(* IEC 61131-3 sources: station-control-three-platforms/codesys/src (part 2) *)

(* ---- GVL_TestResult.st ---- *)
// Result of the test bench (FB_TestBench). Port of DB_TestResult; read by codesys/scripts/build_and_run.py.
{attribute 'qualified_only'}
VAR_GLOBAL
    Done : BOOL;   // the bench has finished; the values below no longer change
    AllPassed : BOOL;   // Done and every case passed
    CasesTotal : INT;
    CasesRun : INT;
    CasesPassed : INT;
    CasesFailed : INT;
    FirstFailedCase : INT;   // 0 = none
    FirstFailedCheck : INT;   // 0 = none; codes in the header of FB_TestBench
    MaxFeatError : REAL;   // N or mm, largest difference of an element from its expected value
    BenchCalls : DINT;   // task cycles the bench needed
    CasePass : ARRAY[1..32] OF BOOL;
    CaseCheck : ARRAY[1..32] OF INT;   // failed check of each case, 0 = passed
    CaseNok : ARRAY[1..32] OF INT;   // NOK code the block gave in each case
END_VAR

(* ---- FB_CurveEval.st ---- *)
FUNCTION_BLOCK FB_CurveEval
//  CODESYS V3.5 port of the Siemens SCL block. Only the syntax changed: no # before local names,
//  REGION as {region} pragma, global data as qualified GVL names, LIMIT with positional arguments.
//  Called in the cyclic interrupt that samples the load cell and the axis position.
//  Nothing is stored as a curve: every evaluation element is updated with the new sample.
//  The block works on static variables and writes its outputs once, at the end of every call.
//  Elements (DOSSIER section 6.3):
//    gate 1 (GateX)    pull force FpG1 and return force FrG1 at the same travel;
//                      FMean = (FpG1 + FrG1) / 2 is the spring, FHyst = FpG1 - FrG1 is twice the friction
//    gate 2 (Gate2X)   pull force after the cable is taut
//    peak window       highest pull force between PeakXLo and PeakXHi and its travel (latch release)
//    step              force drop within StepSpan after the peak
//    stop              travel at which the pull force crosses StopF (end stop)
//    envelope          pull force at fixed travel nodes against EnvLo / EnvHi
//  Mode: 1 peak force only, 2 pull-stroke windows, 3 windows with return stroke, 4 envelope.
//  NokCode: 0 OK, 1 element not measured, 2 gate-1 force (spring), 3 hysteresis (friction),
//           4 no return force, 5 gate-2 force, 6 peak force, 7 peak travel, 8 release step,
//           9 stop travel, 10 envelope.
   VAR_INPUT
      Reset : Bool;   // clear all results, before a new pull
      Sample : Bool;   // X and F are a new sample
      Stroke : Int;   // 1 pull, 2 return
      X : Real;   // mm, travel from touch
      F : Real;   // N
      Finish : Bool;   // return stroke finished: judge
      Mode : Int := 3;
      GateX : Real := 3.0;   // mm
      Gate2X : Real := 10.0;   // mm
      PeakXLo : Real := 13.0;   // mm
      PeakXHi : Real := 26.0;   // mm
      StepSpan : Real := 2.0;   // mm
      StopF : Real := 30.0;   // N
      G1Lo : Real;   // N, limits of FpG1 (mode 2)
      G1Hi : Real;
      MeanLo : Real;   // N, limits of FMean (mode 3)
      MeanHi : Real;
      HystLo : Real;   // N, limits of FHyst (mode 3)
      HystHi : Real;
      RetFMin : Real;   // N, FrG1 must be above (mode 3)
      G2Lo : Real;   // N, limits of FpG2
      G2Hi : Real;
      PeakFLo : Real;   // N
      PeakFHi : Real;
      PeakXMin : Real;   // mm, limits of XPeak
      PeakXMax : Real;
      StepLo : Real;   // N
      StopXLo : Real;   // mm
      StopXHi : Real;
      EnvX0 : Real := 1.0;   // mm, first envelope node
      EnvDx : Real := 0.5;   // mm, node spacing
      EnvN : Int := 55;   // number of nodes, at most 64
      EnvLo : Array[0..63] of Real;   // N
      EnvHi : Array[0..63] of Real;   // N
   END_VAR

   VAR_OUTPUT
      FpG1 : Real;
      FrG1 : Real;
      FMean : Real;
      FHyst : Real;
      FpG2 : Real;
      FPeak : Real;
      XPeak : Real;
      FStep : Real;
      XStop : Real;
      EnvViol : Int;   // envelope nodes outside the band
      EnvNodes : Int;   // envelope nodes evaluated
      NSamples : Int;
      Done : Bool;
      Ok : Bool;
      NokCode : Int;
   END_VAR

   VAR
      sHavePrev : Bool;
      sPrevX : Real;
      sPrevF : Real;
      sPrevStroke : Int;
      sGotG1 : Bool;
      sGotG2 : Bool;
      sGotR1 : Bool;
      sGotPeak : Bool;
      sGotStop : Bool;
      sFMin : Real;
      sFpG1 : Real;
      sFrG1 : Real;
      sFMean : Real;
      sFHyst : Real;
      sFpG2 : Real;
      sFPeak : Real;
      sXPeak : Real;
      sFStep : Real;
      sXStop : Real;
      sEnvViol : Int;
      sEnvNodes : Int;
      sNSamples : Int;
      sDone : Bool;
      sOk : Bool;
      sNokCode : Int;
   END_VAR

   VAR_TEMP
      tI : Int;
      tNodeX : Real;
      tFn : Real;
      tCode : Int;
   END_VAR

(* @IMPLEMENTATION *)
    {region "Reset"}
        IF Reset THEN
            sFpG1 := 0.0;
            sFrG1 := 0.0;
            sFMean := 0.0;
            sFHyst := 0.0;
            sFpG2 := 0.0;
            sFPeak := 0.0;
            sXPeak := 0.0;
            sFStep := 0.0;
            sXStop := 0.0;
            sEnvViol := 0;
            sEnvNodes := 0;
            sNSamples := 0;
            sDone := FALSE;
            sOk := FALSE;
            sNokCode := 0;
            sHavePrev := FALSE;
            sGotG1 := FALSE;
            sGotG2 := FALSE;
            sGotR1 := FALSE;
            sGotPeak := FALSE;
            sGotStop := FALSE;
            sFMin := 0.0;
        END_IF;
    {endregion}

    {region "PullStroke"}
        IF NOT Reset AND Sample AND NOT sDone AND Stroke = 1 THEN
            IF sHavePrev AND sPrevStroke = 1 THEN
                // gates: force at a set travel, linear between the two samples around it
                IF NOT sGotG1 AND sPrevX < GateX AND X >= GateX THEN
                    sFpG1 := sPrevF + (F - sPrevF) * (GateX - sPrevX) / (X - sPrevX);
                    sGotG1 := TRUE;
                END_IF;
                IF NOT sGotG2 AND sPrevX < Gate2X AND X >= Gate2X THEN
                    sFpG2 := sPrevF + (F - sPrevF) * (Gate2X - sPrevX) / (X - sPrevX);
                    sGotG2 := TRUE;
                END_IF;
                // end stop: travel at a set force
                IF NOT sGotStop AND sPrevX > Gate2X AND sPrevF < StopF AND F >= StopF THEN
                    sXStop := sPrevX + (X - sPrevX) * (StopF - sPrevF) / (F - sPrevF);
                    sGotStop := TRUE;
                END_IF;
                // envelope: at most four nodes can lie between two samples
                FOR tI := 1 TO 4 DO
                    tNodeX := EnvX0 + EnvDx * INT_TO_REAL(sEnvNodes);
                    IF sEnvNodes < EnvN AND sPrevX < tNodeX AND X >= tNodeX THEN
                        tFn := sPrevF + (F - sPrevF) * (tNodeX - sPrevX) / (X - sPrevX);
                        IF tFn < EnvLo[sEnvNodes] OR tFn > EnvHi[sEnvNodes] THEN
                            sEnvViol := sEnvViol + 1;
                        END_IF;
                        sEnvNodes := sEnvNodes + 1;
                    END_IF;
                END_FOR;
            END_IF;
            // latch release: peak inside the window, then the drop after it
            IF X >= PeakXLo AND X <= PeakXHi AND (NOT sGotPeak OR F > sFPeak) THEN
                sFPeak := F;
                sXPeak := X;
                sFMin := F;
                sGotPeak := TRUE;
            ELSIF sGotPeak AND X <= sXPeak + StepSpan AND F < sFMin THEN
                sFMin := F;
            END_IF;
            IF sGotPeak THEN
                sFStep := sFPeak - sFMin;
            END_IF;
        END_IF;
    {endregion}

    {region "ReturnStroke"}
        IF NOT Reset AND Sample AND NOT sDone AND Stroke = 2 AND sHavePrev THEN
            IF NOT sGotR1 AND sPrevX > GateX AND X <= GateX THEN
                sFrG1 := sPrevF + (F - sPrevF) * (GateX - sPrevX) / (X - sPrevX);
                sGotR1 := TRUE;
            END_IF;
        END_IF;
    {endregion}

    {region "Bookkeeping"}
        IF NOT Reset AND Sample AND NOT sDone THEN
            sPrevX := X;
            sPrevF := F;
            sPrevStroke := Stroke;
            sHavePrev := TRUE;
            IF sNSamples < 32000 THEN
                sNSamples := sNSamples + 1;
            END_IF;
        END_IF;
    {endregion}

    {region "Verdict"}
        IF NOT Reset AND Finish AND NOT sDone THEN
            sFMean := (sFpG1 + sFrG1) * 0.5;
            sFHyst := sFpG1 - sFrG1;
            tCode := 0;
            CASE Mode OF
                1:  // peak force only
                    IF NOT sGotPeak THEN
                        tCode := 1;
                    ELSIF sFPeak < PeakFLo OR sFPeak > PeakFHi THEN
                        tCode := 6;
                    END_IF;
                2, 3:  // windows; mode 3 judges gate 1 with the return stroke
                    IF NOT (sGotG1 AND sGotG2 AND sGotPeak AND sGotStop) THEN
                        tCode := 1;
                    ELSIF Mode = 3 AND NOT sGotR1 THEN
                        tCode := 1;
                    ELSIF Mode = 2 AND (sFpG1 < G1Lo OR sFpG1 > G1Hi) THEN
                        tCode := 2;
                    ELSIF Mode = 3 AND (sFMean < MeanLo OR sFMean > MeanHi) THEN
                        tCode := 2;
                    ELSIF Mode = 3 AND (sFHyst < HystLo OR sFHyst > HystHi) THEN
                        tCode := 3;
                    ELSIF Mode = 3 AND sFrG1 < RetFMin THEN
                        tCode := 4;
                    ELSIF sFpG2 < G2Lo OR sFpG2 > G2Hi THEN
                        tCode := 5;
                    ELSIF sFPeak < PeakFLo OR sFPeak > PeakFHi THEN
                        tCode := 6;
                    ELSIF sXPeak < PeakXMin OR sXPeak > PeakXMax THEN
                        tCode := 7;
                    ELSIF sFStep < StepLo THEN
                        tCode := 8;
                    ELSIF sXStop < StopXLo OR sXStop > StopXHi THEN
                        tCode := 9;
                    END_IF;
                4:  // envelope: every node reached and inside
                    IF sEnvNodes < EnvN THEN
                        tCode := 1;
                    ELSIF sEnvViol > 0 THEN
                        tCode := 10;
                    END_IF;
                ELSE
                    tCode := 1;
            END_CASE;
            sNokCode := tCode;
            sOk := tCode = 0;
            sDone := TRUE;
        END_IF;
    {endregion}

    {region "Outputs"}
        // the working values live in static variables; the outputs are written here and nowhere else
        FpG1 := sFpG1;
        FrG1 := sFrG1;
        FMean := sFMean;
        FHyst := sFHyst;
        FpG2 := sFpG2;
        FPeak := sFPeak;
        XPeak := sXPeak;
        FStep := sFStep;
        XStop := sXStop;
        EnvViol := sEnvViol;
        EnvNodes := sEnvNodes;
        NSamples := sNSamples;
        Done := sDone;
        Ok := sOk;
        NokCode := sNokCode;
    {endregion}
END_FUNCTION_BLOCK

(* ---- FB_HandleStation.st ---- *)
FUNCTION_BLOCK FB_HandleStation
//  CODESYS V3.5 port of the Siemens SCL block (siemens/scl/FB_HandleStation.scl). Changes, all forced
//  by the compiler: the timer variable sT is sTim (ST is a keyword, identifiers are not case-sensitive);
//  the evaluation recipe comes in by reference (Rcp) and is copied into Eval at the tare, because the
//  caller may not write into Eval from outside (C0037).
//  Called in the same cyclic interrupt as the sampling (CycleTime).
//  States (DOSSIER section 3):
//    0 Idle         wait for a part; check presence time and the LH/RH sensor pattern
//    1 Clamp        close the clamp
//    2 Tare         zero the load cell with the hook free
//    3 Approach     drive towards the grip until the force passes FTouch; the touch position
//                   must lie in its window
//    4 Pull         sample every cycle into the curve evaluation; reverse at FRev
//    5 Return       sample the return stroke down to travel 0, then go home fast
//    6 Evaluate     judge
//    7 UnloadOk     open the clamp; wait until the part has left
//    8 RejectLock   open the clamp; the station stays locked until the part has left AND the
//                   reject-chute sensor has seen a part pass
//    9 Fault        drive stopped; after the acknowledge the axis goes home and the part that was
//                   in test is treated as rejected (an interrupted test is not a passed test)
//   10 Home         go home after a fault
//  NokCode: 1 to 10 from FB_CurveEval; 20 wrong hand or sensor pattern not plausible;
//           21 no touch or touch outside its window; 22 force above FAbsMax; 23 no end stop;
//           24 test interrupted by a fault.
//  FaultCode: 1 safety circuit open, 2 drive not ready, 3 clamp time-out, 4 load cell does not tare.
   VAR_INPUT
      CycleTime : Real := 0.002;   // s
      SafetyOk : Bool;
      DriveOk : Bool;
      AckFault : Bool;
      StartEnable : Bool;   // release from the line
      PartPresent : Bool;
      SensLH : Bool;   // variant sensor that only an LH unit covers
      SensRH : Bool;   // variant sensor that only an RH unit covers
      VariantLH : Bool;   // recipe: TRUE = LH units are being built
      ClampClosed : Bool;
      ClampOpen : Bool;
      RejectChute : Bool;   // light barrier in the reject chute
      Pos : Real;   // mm, axis position, 0 = home
      Force : Real;   // N, load cell
      VPull : Real := 50.0;   // mm/s
      VHome : Real := 150.0;   // mm/s
      FTouch : Real := 1.5;   // N
      FRev : Real := 40.0;   // N
      FAbsMax : Real := 60.0;   // N, protects the painted part
      XMax : Real := 38.0;   // mm
      TouchLo : Real := 3.0;   // mm, window of the touch position
      TouchHi : Real := 7.0;
      Compliance : Real := 0.025;   // mm/N, rig deflection taken out of the travel
      TareTol : Real := 0.5;   // N
      TPresent : Real := 0.1;   // s
      TClampMax : Real := 1.0;   // s
      TRejectWarn : Real := 30.0;   // s
      MaxConsecNok : Int := 3;
   END_VAR

   VAR_IN_OUT
      Rcp : ST_EvalRecipe;   // evaluation recipe, copied into Eval at every tare
   END_VAR

   VAR_OUTPUT
      QClamp : Bool;
      QDriveEnable : Bool;
      QVel : Real;   // mm/s, positive = pull
      QLampOk : Bool;
      QLampNok : Bool;
      QCallOperator : Bool;
      State : Int;
      Verdict : Int;   // 0 none, 1 OK, 2 NOK
      NokCode : Int;
      FaultCode : Int;
      Locked : Bool;
      RigCheckRequired : Bool;   // too many rejects in a row: run the master part
      XTravel : Real;   // mm
      FNet : Real;   // N
      TCycle : Real;   // s, clamp to verdict of the last part
      CntTotal : DInt;
      CntOk : DInt;
      CntNok : DInt;
      CntRejectConfirmed : DInt;
      CntConsecNok : Int;
      CntByCode : Array[0..31] of DInt;
   END_VAR

   VAR
      Eval : FB_CurveEval;
      sTim : Real;
      sTCycle : Real;
      sTare : Real;
      sTouchPos : Real;
      sFTouch : Real;
      sPreNok : Int;
      sPartGone : Bool;
      sChutePrev : Bool;
      sInTest : Bool;
      sWasLocked : Bool;
      sState : Int;
      sRigCheckRequired : Bool;
      sCntTotal : DInt;
      sCntOk : DInt;
      sCntNok : DInt;
      sCntRejectConfirmed : DInt;
      sCntConsecNok : Int;
      sCntByCode : Array[0..31] of DInt;
   END_VAR

   VAR_TEMP
      tVariantOk : Bool;
      tChuteEdge : Bool;
      tCode : Int;
   END_VAR

(* @IMPLEMENTATION *)
    {region "Inputs"}
        FNet := Force - sTare;
        tChuteEdge := RejectChute AND NOT sChutePrev;
        sChutePrev := RejectChute;
        sTim := sTim + CycleTime;
        sTCycle := sTCycle + CycleTime;
        QVel := 0.0;
        // exactly the sensor of the expected hand, and not the other one
        tVariantOk := (VariantLH AND SensLH AND NOT SensRH) OR (NOT VariantLH AND SensRH AND NOT SensLH);
    {endregion}

    {region "Faults"}
        IF sState <> 9 AND (NOT SafetyOk OR NOT DriveOk) THEN
            IF NOT SafetyOk THEN
                FaultCode := 1;
            ELSE
                FaultCode := 2;
            END_IF;
            IF sState <> 10 THEN
                sInTest := sState >= 1 AND sState <= 6;
                sWasLocked := sState = 8;
            END_IF;
            sState := 9;
        END_IF;
    {endregion}

    {region "Sequence"}
        CASE sState OF
            0:  // Idle
                Locked := FALSE;
                IF NOT PartPresent THEN
                    sTim := 0.0;
                    QLampOk := FALSE;
                    QLampNok := FALSE;
                ELSIF sTim >= TPresent AND StartEnable AND ClampOpen AND NOT sRigCheckRequired THEN
                    Verdict := 0;
                    NokCode := 0;
                    sPreNok := 0;
                    sTCycle := 0.0;
                    sTim := 0.0;
                    IF tVariantOk THEN
                        sState := 1;
                    ELSE
                        sPreNok := 20;   // never pull a part of the wrong hand
                        sState := 6;
                    END_IF;
                END_IF;
            1:  // Clamp
                QClamp := TRUE;
                IF ClampClosed THEN
                    sTim := 0.0;
                    sState := 2;
                ELSIF sTim > TClampMax THEN
                    FaultCode := 3;
                    sInTest := TRUE;
                    sState := 9;
                END_IF;
            2:  // Tare
                IF sTim >= 0.05 THEN
                    IF ABS(Force) > TareTol THEN
                        FaultCode := 4;
                        sInTest := TRUE;
                        sState := 9;
                    ELSE
                        sTare := Force;
                        // the recipe of this part (Siemens: written into Eval by the caller)
                        Eval.Mode := Rcp.Mode;
                        Eval.GateX := Rcp.GateX;
                        Eval.Gate2X := Rcp.Gate2X;
                        Eval.PeakXLo := Rcp.PeakXLo;
                        Eval.PeakXHi := Rcp.PeakXHi;
                        Eval.StepSpan := Rcp.StepSpan;
                        Eval.StopF := Rcp.StopF;
                        Eval.G1Lo := Rcp.G1Lo;
                        Eval.G1Hi := Rcp.G1Hi;
                        Eval.MeanLo := Rcp.MeanLo;
                        Eval.MeanHi := Rcp.MeanHi;
                        Eval.HystLo := Rcp.HystLo;
                        Eval.HystHi := Rcp.HystHi;
                        Eval.RetFMin := Rcp.RetFMin;
                        Eval.G2Lo := Rcp.G2Lo;
                        Eval.G2Hi := Rcp.G2Hi;
                        Eval.PeakFLo := Rcp.PeakFLo;
                        Eval.PeakFHi := Rcp.PeakFHi;
                        Eval.PeakXMin := Rcp.PeakXMin;
                        Eval.PeakXMax := Rcp.PeakXMax;
                        Eval.StepLo := Rcp.StepLo;
                        Eval.StopXLo := Rcp.StopXLo;
                        Eval.StopXHi := Rcp.StopXHi;
                        Eval.EnvX0 := Rcp.EnvX0;
                        Eval.EnvDx := Rcp.EnvDx;
                        Eval.EnvN := Rcp.EnvN;
                        Eval.EnvLo := Rcp.EnvLo;
                        Eval.EnvHi := Rcp.EnvHi;
                        Eval(Reset := TRUE, Sample := FALSE, Stroke := 0, X := 0.0, F := 0.0, Finish := FALSE);
                        sState := 3;
                    END_IF;
                END_IF;
            3:  // Approach
                QVel := VPull;
                IF FNet > FTouch THEN
                    sTouchPos := Pos;
                    sFTouch := FNet;
                    IF Pos < TouchLo OR Pos > TouchHi THEN
                        sPreNok := 21;
                        sState := 5;
                    ELSE
                        XTravel := 0.0;
                        Eval(Reset := FALSE, Sample := TRUE, Stroke := 1, X := 0.0, F := FNet, Finish := FALSE);
                        sState := 4;
                    END_IF;
                ELSIF Pos > TouchHi THEN
                    sPreNok := 21;
                    sTouchPos := Pos;
                    sFTouch := 0.0;
                    sState := 5;
                END_IF;
            4:  // Pull
                QVel := VPull;
                XTravel := Pos - sTouchPos - (FNet - sFTouch) * Compliance;
                Eval(Reset := FALSE, Sample := TRUE, Stroke := 1, X := XTravel, F := FNet, Finish := FALSE);
                IF FNet >= FAbsMax THEN
                    sPreNok := 22;
                    sState := 5;
                ELSIF FNet >= FRev THEN
                    sState := 5;
                ELSIF XTravel >= XMax THEN
                    sPreNok := 23;
                    sState := 5;
                END_IF;
            5:  // Return
                XTravel := Pos - sTouchPos - (FNet - sFTouch) * Compliance;
                IF Pos > sTouchPos - 0.5 THEN
                    QVel := -VPull;
                    IF sPreNok = 0 THEN
                        Eval(Reset := FALSE, Sample := TRUE, Stroke := 2, X := XTravel, F := FNet, Finish := FALSE);
                    END_IF;
                ELSIF Pos > 0.05 THEN
                    QVel := -VHome;
                ELSE
                    sState := 6;
                END_IF;
            6:  // Evaluate
                IF sPreNok <> 0 THEN
                    tCode := sPreNok;
                ELSE
                    Eval(Reset := FALSE, Sample := FALSE, Stroke := 0, X := 0.0, F := 0.0, Finish := TRUE);
                    tCode := Eval.NokCode;
                END_IF;
                NokCode := tCode;
                TCycle := sTCycle;
                sCntTotal := sCntTotal + 1;
                sCntByCode[tCode] := sCntByCode[tCode] + 1;
                QClamp := FALSE;
                sTim := 0.0;
                IF tCode = 0 THEN
                    Verdict := 1;
                    sCntOk := sCntOk + 1;
                    sCntConsecNok := 0;
                    QLampOk := TRUE;
                    sState := 7;
                ELSE
                    Verdict := 2;
                    sCntNok := sCntNok + 1;
                    sCntConsecNok := sCntConsecNok + 1;
                    QLampNok := TRUE;
                    sPartGone := FALSE;
                    sState := 8;
                END_IF;
            7:  // UnloadOk
                QClamp := FALSE;
                IF NOT PartPresent AND ClampOpen THEN
                    sTim := 0.0;
                    sState := 0;
                END_IF;
            8:  // RejectLock
                QClamp := FALSE;
                Locked := TRUE;
                IF NOT PartPresent THEN
                    sPartGone := TRUE;
                END_IF;
                QCallOperator := sTim > TRejectWarn OR sRigCheckRequired;
                IF sPartGone AND tChuteEdge THEN
                    sCntRejectConfirmed := sCntRejectConfirmed + 1;
                    sRigCheckRequired := sCntConsecNok >= MaxConsecNok;
                    QCallOperator := sRigCheckRequired;
                    Locked := FALSE;
                    sTim := 0.0;
                    sState := 0;
                END_IF;
            9:  // Fault
                QClamp := sInTest;
                QCallOperator := TRUE;
                IF AckFault AND SafetyOk AND DriveOk THEN
                    FaultCode := 0;
                    QCallOperator := FALSE;
                    sState := 10;
                END_IF;
            10:  // Home
                IF Pos > 0.05 THEN
                    QVel := -VPull;
                ELSIF sInTest THEN
                    sInTest := FALSE;
                    sPreNok := 24;
                    sState := 6;
                ELSIF sWasLocked THEN
                    sWasLocked := FALSE;   // a fault does not release the reject lock
                    sState := 8;
                ELSE
                    sState := 0;
                END_IF;
            ELSE
                sState := 9;
        END_CASE;
    {endregion}

    {region "RigCheck"}
        // the lock after too many rejects in a row is released by the acknowledge key
        IF sRigCheckRequired AND AckFault AND sState = 0 THEN
            sRigCheckRequired := FALSE;
            sCntConsecNok := 0;
            QCallOperator := FALSE;
        END_IF;
        QDriveEnable := SafetyOk AND DriveOk AND sState <> 9;
    {endregion}

    {region "Outputs"}
        // state and counters live in static variables; these outputs are written here and nowhere else
        State := sState;
        RigCheckRequired := sRigCheckRequired;
        CntTotal := sCntTotal;
        CntOk := sCntOk;
        CntNok := sCntNok;
        CntRejectConfirmed := sCntRejectConfirmed;
        CntConsecNok := sCntConsecNok;
        CntByCode := sCntByCode;
    {endregion}
END_FUNCTION_BLOCK

(* ---- FB_TestBench.st ---- *)
FUNCTION_BLOCK FB_TestBench
//  CODESYS V3.5 port of siemens/scl/test/FB_TestBench.scl. Changes: sT is sTim; the station recipe is
//  the local structure StationRcp, passed to the station as Rcp (Siemens: Station.Eval.* written directly).
//  Called from OB1 every cycle. Needs no input from outside. Finishes on its own, then holds its
//  result in DB_TestResult.
//  Part 1, replay cases 1..NCases (DB_TestData): a recorded curve goes sample by sample into
//    FB_CurveEval. Verdict, NOK code, the nine elements and the envelope counts must equal the
//    values the NumPy evaluation gave for the same samples (elements within DB_TestData.Tol).
//  Part 2, six station cases: FB_HandleStation runs against FB_TestPlant.
//    NCases+1  good LH unit is clamped, pulled and passed
//    NCases+2  RH unit on an LH recipe: reject code 20, axis and clamp never move
//    NCases+3  reject lock: a chute signal while the part is in the fixture does not open it, a new
//              part is not started, the chute signal after the fixture is empty opens it
//    NCases+4  unit with unhooked latch lever: pulled, reject code 5
//    NCases+5  third reject in a row: master part asked for, start blocked
//    NCases+6  after the acknowledge the good unit is pulled and passed
//  Check codes (DB_TestResult.FirstFailedCheck, CaseCheck): 0 passed.
//    Replay:  1 verdict, 2 NOK code, 3 FpG1, 4 FrG1, 5 FMean, 6 FHyst, 7 FpG2, 8 FPeak, 9 XPeak,
//             10 FStep, 11 XStop, 12 envelope nodes outside, 13 envelope nodes evaluated
//    Station: 21 verdict, 22 NOK code, 23 state, 24 counter, 25 axis or clamp moved (or did not),
//             26 reject lock opened too early or a part was started while locked,
//             27 reject lock not opened by the chute, 28 master-part request, 29 time-out
   VAR_INPUT
      ReplayPerCall : Int := 200;   // samples replayed per call
      ScansPerCall : Int := 100;   // station scans (2 ms of station time each) per call
   END_VAR

   VAR
      Eval : FB_CurveEval;
      Station : FB_HandleStation;
      Plant : FB_TestPlant;
      StationRcp : ST_EvalRecipe;   // recipe of the station (Siemens: written into Station.Eval)
      sPhase : Int;   // 0 start, 1 replay, 2 station, 3 done
      sSub : Int;
      sCase : Int;
      sIdx : Int;
      sCk : Int;
      sNok : Int;
      sRecord : Bool;
      sRun : Int;
      sPassed : Int;
      sFailed : Int;
      sFirstCase : Int;
      sFirstCheck : Int;
      sMaxErr : Real;
      sCalls : DInt;
      sMeas : Array[0..8] of Real;
      sStep : Int;
      sTim : Int;
      sPart : Bool;
      sLH : Bool;
      sRH : Bool;
      sChute : Bool;
      sAck : Bool;
      sPlantReset : Bool;
      sCurve : Int;
   END_VAR

   VAR_TEMP
      tI : Int;
      tJ : Int;
      tB : Int;
      tCurve : Int;
      tMode : Int;
      tA : Int;
      tN : Int;
      tStroke : Int;
      tErr : Real;
   END_VAR

(* @IMPLEMENTATION *)
    {region "Start"}
        IF sPhase = 0 THEN
            FOR tI := 1 TO 32 DO
                GVL_TestResult.CasePass[tI] := FALSE;
                GVL_TestResult.CaseCheck[tI] := 0;
                GVL_TestResult.CaseNok[tI] := 0;
            END_FOR;
            // the part of the recipe that is the same in every case, for both evaluation instances
            Eval.GateX := GVL_TestData.GateX;
            Eval.Gate2X := GVL_TestData.Gate2X;
            Eval.PeakXLo := GVL_TestData.PeakXLo;
            Eval.PeakXHi := GVL_TestData.PeakXHi;
            Eval.StepSpan := GVL_TestData.StepSpan;
            Eval.StopF := GVL_TestData.StopF;
            Eval.EnvX0 := GVL_TestData.EnvX0;
            Eval.EnvDx := GVL_TestData.EnvDx;
            Eval.EnvN := GVL_TestData.EnvN;
            StationRcp.GateX := GVL_TestData.GateX;
            StationRcp.Gate2X := GVL_TestData.Gate2X;
            StationRcp.PeakXLo := GVL_TestData.PeakXLo;
            StationRcp.PeakXHi := GVL_TestData.PeakXHi;
            StationRcp.StepSpan := GVL_TestData.StepSpan;
            StationRcp.StopF := GVL_TestData.StopF;
            StationRcp.EnvX0 := GVL_TestData.EnvX0;
            StationRcp.EnvDx := GVL_TestData.EnvDx;
            StationRcp.EnvN := GVL_TestData.EnvN;
            FOR tI := 0 TO 63 DO
                Eval.EnvLo[tI] := GVL_TestData.EnvLo[tI];
                Eval.EnvHi[tI] := GVL_TestData.EnvHi[tI];
                StationRcp.EnvLo[tI] := GVL_TestData.EnvLo[tI];
                StationRcp.EnvHi[tI] := GVL_TestData.EnvHi[tI];
            END_FOR;
            // the station judges with windows + return stroke (mode 3: limits 32..47)
            StationRcp.Mode := 3;
            StationRcp.G1Lo := GVL_TestData.Lim[32];
            StationRcp.G1Hi := GVL_TestData.Lim[33];
            StationRcp.MeanLo := GVL_TestData.Lim[34];
            StationRcp.MeanHi := GVL_TestData.Lim[35];
            StationRcp.HystLo := GVL_TestData.Lim[36];
            StationRcp.HystHi := GVL_TestData.Lim[37];
            StationRcp.RetFMin := GVL_TestData.Lim[38];
            StationRcp.G2Lo := GVL_TestData.Lim[39];
            StationRcp.G2Hi := GVL_TestData.Lim[40];
            StationRcp.PeakFLo := GVL_TestData.Lim[41];
            StationRcp.PeakFHi := GVL_TestData.Lim[42];
            StationRcp.PeakXMin := GVL_TestData.Lim[43];
            StationRcp.PeakXMax := GVL_TestData.Lim[44];
            StationRcp.StepLo := GVL_TestData.Lim[45];
            StationRcp.StopXLo := GVL_TestData.Lim[46];
            StationRcp.StopXHi := GVL_TestData.Lim[47];
            sCase := 1;
            sSub := 0;
            sCk := 0;
            sNok := 0;
            sStep := 10;
            sTim := 0;
            sPhase := 1;
        END_IF;
        IF sPhase < 3 THEN
            sCalls := sCalls + 1;
        END_IF;
    {endregion}

    {region "Replay"}
        IF sPhase = 1 THEN
            FOR tI := 1 TO ReplayPerCall DO
                IF NOT sRecord THEN
                    tCurve := GVL_TestData.CaseCurve[sCase];
                    tMode := GVL_TestData.CaseMode[sCase];
                    tA := GVL_TestData.CurveStart[tCurve];
                    tN := GVL_TestData.CurveNPull[tCurve];
                    CASE sSub OF
                        0:  // limits of the mode of this case, clear the evaluation
                            tB := (tMode - 1) * 16;
                            Eval.Mode := tMode;
                            Eval.G1Lo := GVL_TestData.Lim[tB];
                            Eval.G1Hi := GVL_TestData.Lim[tB + 1];
                            Eval.MeanLo := GVL_TestData.Lim[tB + 2];
                            Eval.MeanHi := GVL_TestData.Lim[tB + 3];
                            Eval.HystLo := GVL_TestData.Lim[tB + 4];
                            Eval.HystHi := GVL_TestData.Lim[tB + 5];
                            Eval.RetFMin := GVL_TestData.Lim[tB + 6];
                            Eval.G2Lo := GVL_TestData.Lim[tB + 7];
                            Eval.G2Hi := GVL_TestData.Lim[tB + 8];
                            Eval.PeakFLo := GVL_TestData.Lim[tB + 9];
                            Eval.PeakFHi := GVL_TestData.Lim[tB + 10];
                            Eval.PeakXMin := GVL_TestData.Lim[tB + 11];
                            Eval.PeakXMax := GVL_TestData.Lim[tB + 12];
                            Eval.StepLo := GVL_TestData.Lim[tB + 13];
                            Eval.StopXLo := GVL_TestData.Lim[tB + 14];
                            Eval.StopXHi := GVL_TestData.Lim[tB + 15];
                            Eval(Reset := TRUE, Sample := FALSE, Stroke := 0, X := 0.0, F := 0.0, Finish := FALSE);
                            sIdx := 0;
                            sSub := 1;
                        1:  // one sample: the pull samples first, then the return samples
                            IF sIdx < tN THEN
                                tStroke := 1;
                            ELSE
                                tStroke := 2;
                            END_IF;
                            Eval(Reset := FALSE, Sample := TRUE, Stroke := tStroke,
                                  X := GVL_TestData.X[tA + sIdx], F := GVL_TestData.F[tA + sIdx], Finish := FALSE);
                            sIdx := sIdx + 1;
                            IF sIdx >= 2 * tN THEN
                                sSub := 2;
                            END_IF;
                        2:  // judge and compare with the expected values
                            Eval(Reset := FALSE, Sample := FALSE, Stroke := 0, X := 0.0, F := 0.0, Finish := TRUE);
                            sMeas[0] := Eval.FpG1;
                            sMeas[1] := Eval.FrG1;
                            sMeas[2] := Eval.FMean;
                            sMeas[3] := Eval.FHyst;
                            sMeas[4] := Eval.FpG2;
                            sMeas[5] := Eval.FPeak;
                            sMeas[6] := Eval.XPeak;
                            sMeas[7] := Eval.FStep;
                            sMeas[8] := Eval.XStop;
                            IF Eval.Ok XOR GVL_TestData.ExpOk[sCase] THEN
                                sCk := 1;
                            ELSIF Eval.NokCode <> GVL_TestData.ExpNok[sCase] THEN
                                sCk := 2;
                            ELSIF Eval.EnvViol <> GVL_TestData.ExpEnvViol[sCase] THEN
                                sCk := 12;
                            ELSIF Eval.EnvNodes <> GVL_TestData.ExpEnvNodes[sCase] THEN
                                sCk := 13;
                            END_IF;
                            FOR tJ := 0 TO 8 DO
                                tB := (sCase - 1) * 9 + tJ;
                                IF GVL_TestData.ExpFeatValid[tB] THEN
                                    tErr := ABS(sMeas[tJ] - GVL_TestData.ExpFeat[tB]);
                                    IF tErr > sMaxErr THEN
                                        sMaxErr := tErr;
                                    END_IF;
                                    IF tErr > GVL_TestData.Tol AND sCk = 0 THEN
                                        sCk := 3 + tJ;
                                    END_IF;
                                END_IF;
                            END_FOR;
                            sNok := Eval.NokCode;
                            sSub := 0;
                            sRecord := TRUE;
                    END_CASE;
                END_IF;
            END_FOR;
        END_IF;
    {endregion}

    {region "Station"}
        IF sPhase = 2 THEN
            FOR tI := 1 TO ScansPerCall DO
                IF sPhase = 2 AND NOT sRecord THEN
                    IF sTim < 30000 THEN
                        sTim := sTim + 1;
                    END_IF;
                    // what the operator and the line do, and what the station must have done by now
                    CASE sStep OF
                        10:  // good LH unit
                            sPart := TRUE;
                            sLH := TRUE;
                            sRH := FALSE;
                            sCurve := GVL_TestData.GoodCurve;
                            sPlantReset := TRUE;
                            sStep := 11;
                            sTim := 0;
                        11:
                            IF Station.CntTotal >= 1 OR sTim > 4000 THEN
                                IF sTim > 4000 THEN
                                    sCk := 29;
                                ELSIF Station.Verdict <> 1 THEN
                                    sCk := 21;
                                ELSIF Station.NokCode <> 0 THEN
                                    sCk := 22;
                                ELSIF Station.CntOk <> 1 OR Station.CntNok <> 0 THEN
                                    sCk := 24;
                                ELSIF NOT Plant.Moved THEN
                                    sCk := 25;
                                END_IF;
                                sNok := Station.NokCode;
                                sRecord := TRUE;
                                sPart := FALSE;
                                sStep := 12;
                                sTim := 0;
                            END_IF;
                        12:  // unit taken out
                            IF Station.State = 0 OR sTim > 4000 THEN
                                sStep := 20;
                                sTim := 0;
                            END_IF;
                        20:  // RH unit while LH units are built
                            sPart := TRUE;
                            sLH := FALSE;
                            sRH := TRUE;
                            sCurve := GVL_TestData.GoodCurve;
                            sPlantReset := TRUE;
                            sStep := 21;
                            sTim := 0;
                        21:
                            IF Station.CntTotal >= 2 OR sTim > 4000 THEN
                                IF sTim > 4000 THEN
                                    sCk := 29;
                                ELSIF Station.Verdict <> 2 THEN
                                    sCk := 21;
                                ELSIF Station.NokCode <> 20 THEN
                                    sCk := 22;
                                ELSIF Station.State <> 8 THEN
                                    sCk := 23;
                                ELSIF Plant.Moved OR Plant.Pos > 0.0 OR NOT Plant.ClampOpen THEN
                                    sCk := 25;
                                END_IF;
                                sNok := Station.NokCode;
                                sRecord := TRUE;
                                sStep := 22;
                                sTim := 0;
                            END_IF;
                        22:  // reject lock: a chute signal while the rejected unit is still in the fixture
                            sChute := sTim >= 5 AND sTim < 10;
                            IF sTim >= 20 THEN
                                IF Station.State <> 8 OR NOT Station.Locked THEN
                                    sCk := 26;
                                END_IF;
                                sPart := FALSE;
                                sStep := 23;
                                sTim := 0;
                            END_IF;
                        23:  // the unit is taken out and a new good unit is put in without using the chute
                            IF sTim = 20 THEN
                                sPart := TRUE;
                                sLH := TRUE;
                                sRH := FALSE;
                                sPlantReset := TRUE;
                            END_IF;
                            IF sTim >= 400 THEN
                                IF sCk = 0 AND (Station.State <> 8 OR Station.CntTotal <> 2 OR Plant.Moved) THEN
                                    sCk := 26;
                                END_IF;
                                sPart := FALSE;
                                sStep := 24;
                                sTim := 0;
                            END_IF;
                        24:  // fixture empty, the chute sensor sees a part
                            sChute := sTim >= 20 AND sTim < 25;
                            IF sTim >= 40 THEN
                                IF sCk = 0 AND (Station.State <> 0 OR Station.Locked OR Station.CntRejectConfirmed <> 1) THEN
                                    sCk := 27;
                                END_IF;
                                sNok := Station.NokCode;
                                sRecord := TRUE;
                                sStep := 30;
                                sTim := 0;
                            END_IF;
                        30:  // LH unit with unhooked latch lever
                            sPart := TRUE;
                            sLH := TRUE;
                            sRH := FALSE;
                            sCurve := GVL_TestData.BadCurve;
                            sPlantReset := TRUE;
                            sStep := 31;
                            sTim := 0;
                        31:
                            IF Station.CntTotal >= 3 OR sTim > 4000 THEN
                                IF sTim > 4000 THEN
                                    sCk := 29;
                                ELSIF Station.Verdict <> 2 THEN
                                    sCk := 21;
                                ELSIF Station.NokCode <> 5 THEN
                                    sCk := 22;
                                ELSIF Station.CntConsecNok <> 2 THEN
                                    sCk := 24;
                                ELSIF NOT Plant.Moved THEN
                                    sCk := 25;
                                END_IF;
                                sNok := Station.NokCode;
                                sRecord := TRUE;
                                sPart := FALSE;
                                sStep := 32;
                                sTim := 0;
                            END_IF;
                        32:  // into the chute
                            sChute := sTim >= 20 AND sTim < 25;
                            IF (sTim >= 40 AND Station.State = 0) OR sTim > 4000 THEN
                                sStep := 40;
                                sTim := 0;
                            END_IF;
                        40:  // the same defect again: third reject in a row
                            sPart := TRUE;
                            sCurve := GVL_TestData.BadCurve;
                            sPlantReset := TRUE;
                            sStep := 41;
                            sTim := 0;
                        41:
                            IF Station.CntTotal >= 4 OR sTim > 4000 THEN
                                IF sTim > 4000 THEN
                                    sCk := 29;
                                ELSIF Station.Verdict <> 2 THEN
                                    sCk := 21;
                                ELSIF Station.NokCode <> 5 THEN
                                    sCk := 22;
                                ELSIF Station.CntConsecNok <> 3 THEN
                                    sCk := 24;
                                END_IF;
                                sNok := Station.NokCode;
                                sPart := FALSE;
                                sStep := 42;
                                sTim := 0;
                            END_IF;
                        42:  // into the chute; then a good unit is put in
                            sChute := sTim >= 20 AND sTim < 25;
                            IF sTim >= 40 THEN
                                IF sCk = 0 AND Station.State <> 0 THEN
                                    sCk := 27;
                                ELSIF sCk = 0 AND (NOT Station.RigCheckRequired OR NOT Station.QCallOperator) THEN
                                    sCk := 28;
                                END_IF;
                                sPart := TRUE;
                                sCurve := GVL_TestData.GoodCurve;
                                sPlantReset := TRUE;
                                sStep := 43;
                                sTim := 0;
                            END_IF;
                        43:  // the start must stay blocked until the acknowledge
                            IF sTim >= 400 THEN
                                IF sCk = 0 AND (Station.State <> 0 OR Station.CntTotal <> 4 OR Plant.Moved) THEN
                                    sCk := 28;
                                END_IF;
                                sRecord := TRUE;
                                sStep := 50;
                                sTim := 0;
                            END_IF;
                        50:  // acknowledge key; the good unit is then tested
                            sAck := sTim < 5;
                            IF Station.CntTotal >= 5 OR sTim > 4000 THEN
                                IF sTim > 4000 THEN
                                    sCk := 29;
                                ELSIF Station.RigCheckRequired THEN
                                    sCk := 28;
                                ELSIF Station.Verdict <> 1 THEN
                                    sCk := 21;
                                ELSIF Station.NokCode <> 0 THEN
                                    sCk := 22;
                                ELSIF Station.CntOk <> 2 OR Station.CntConsecNok <> 0 THEN
                                    sCk := 24;
                                END_IF;
                                sNok := Station.NokCode;
                                sRecord := TRUE;
                                sPart := FALSE;
                                sAck := FALSE;
                                sStep := 51;
                                sTim := 0;
                            END_IF;
                        51:  // unit taken out
                            IF Station.State = 0 OR sTim > 4000 THEN
                                sStep := 99;
                            END_IF;
                        ELSE
                            sPhase := 3;
                    END_CASE;
                    Plant(Reset := sPlantReset, CycleTime := 0.002, QVel := Station.QVel,
                           QDriveEnable := Station.QDriveEnable, QClamp := Station.QClamp,
                           PartPresent := sPart, Curve := sCurve, Seat := 5.0);
                    sPlantReset := FALSE;
                    Station(Rcp := StationRcp, CycleTime := 0.002, SafetyOk := TRUE, DriveOk := TRUE, AckFault := sAck,
                             StartEnable := TRUE, PartPresent := sPart, SensLH := sPart AND sLH,
                             SensRH := sPart AND sRH, VariantLH := TRUE, ClampClosed := Plant.ClampClosed,
                             ClampOpen := Plant.ClampOpen, RejectChute := sChute, Pos := Plant.Pos,
                             Force := Plant.Force, Compliance := 0.0);
                END_IF;
            END_FOR;
        END_IF;
    {endregion}

    {region "Record"}
        IF sRecord THEN
            sRun := sRun + 1;
            IF sCk = 0 THEN
                sPassed := sPassed + 1;
                GVL_TestResult.CasePass[sCase] := TRUE;
            ELSE
                sFailed := sFailed + 1;
                IF sFirstCase = 0 THEN
                    sFirstCase := sCase;
                    sFirstCheck := sCk;
                END_IF;
            END_IF;
            GVL_TestResult.CaseCheck[sCase] := sCk;
            GVL_TestResult.CaseNok[sCase] := sNok;
            sCase := sCase + 1;
            sCk := 0;
            sNok := 0;
            sRecord := FALSE;
            IF sPhase = 1 AND sCase > GVL_TestData.NCases THEN
                sPhase := 2;
            END_IF;
        END_IF;
    {endregion}

    {region "Result"}
        GVL_TestResult.CasesTotal := GVL_TestData.NCases + 6;
        GVL_TestResult.CasesRun := sRun;
        GVL_TestResult.CasesPassed := sPassed;
        GVL_TestResult.CasesFailed := sFailed;
        GVL_TestResult.FirstFailedCase := sFirstCase;
        GVL_TestResult.FirstFailedCheck := sFirstCheck;
        GVL_TestResult.MaxFeatError := sMaxErr;
        GVL_TestResult.BenchCalls := sCalls;
        GVL_TestResult.Done := sPhase = 3;
        GVL_TestResult.AllPassed := sPhase = 3 AND sFailed = 0 AND sPassed = GVL_TestData.NCases + 6;
    {endregion}
END_FUNCTION_BLOCK

(* ---- FB_TestPlant.st ---- *)
FUNCTION_BLOCK FB_TestPlant
//  CODESYS V3.5 port of the Siemens SCL block. Only the syntax changed: no # before local names,
//  REGION as {region} pragma, global data as qualified GVL names, LIMIT with positional arguments.
//  Not part of the station program. Used by FB_TestBench so that FB_HandleStation can run in the
//  PLC without hardware.
//    axis     position follows the speed command, no dynamics
//    clamp    closed 0.25 s after the command, open 0.25 s after it is taken away
//    handle   force read from a recorded curve in DB_TestData at the travel Pos - Seat:
//             the pull samples until the speed command turns negative, the return samples after
//             that; linear between samples; past the last pull sample the end stop goes on at
//             25 N/mm. The recorded travel has the rig deflection taken out already, so the
//             station is run with Compliance = 0.
   VAR_INPUT
      Reset : Bool;   // a new part is in the fixture
      CycleTime : Real := 0.002;   // s
      QVel : Real;   // mm/s
      QDriveEnable : Bool;
      QClamp : Bool;
      PartPresent : Bool;
      Curve : Int;   // recorded curve the part follows
      Seat : Real := 5.0;   // mm, axis position at which the hook meets the grip
   END_VAR

   VAR_OUTPUT
      Pos : Real;   // mm
      Force : Real;   // N
      ClampClosed : Bool;
      ClampOpen : Bool;
      Moved : Bool;   // the axis has moved or the clamp has closed since the last Reset
   END_VAR

   VAR
      sPos : Real;
      sClamp : Real;
      sReturn : Bool;
      sK : Int;
      sMoved : Bool;
   END_VAR

   VAR_TEMP
      tI : Int;
      tA : Int;
      tN : Int;
      tX : Real;
      tF : Real;
      tX0 : Real;
      tX1 : Real;
      tF0 : Real;
      tF1 : Real;
   END_VAR

(* @IMPLEMENTATION *)
    {region "Part"}
        IF Reset THEN
            sReturn := FALSE;
            sK := 0;
            sMoved := FALSE;
        END_IF;
    {endregion}

    {region "AxisAndClamp"}
        IF QDriveEnable THEN
            sPos := sPos + QVel * CycleTime;
            IF QVel <> 0.0 THEN
                sMoved := TRUE;
            END_IF;
        END_IF;
        IF sPos < 0.0 THEN
            sPos := 0.0;
        END_IF;
        IF QClamp THEN
            sClamp := sClamp + CycleTime;
            sMoved := TRUE;
        ELSE
            sClamp := sClamp - CycleTime;
        END_IF;
        sClamp := LIMIT(0.0, sClamp, 0.25);
    {endregion}

    {region "Handle"}
        tX := sPos - Seat;
        tF := 0.0;
        tA := GVL_TestData.CurveStart[Curve];
        tN := GVL_TestData.CurveNPull[Curve];
        IF QVel < 0.0 AND NOT sReturn THEN
            sReturn := TRUE;
            sK := 0;
        END_IF;
        IF PartPresent AND tX >= 0.0 AND tN >= 2 THEN
            IF sReturn THEN
                tA := tA + tN;   // the return samples follow the pull samples; their travel falls
            END_IF;
            // move on to the pair of samples around the travel (the axis moves less than 8 samples per call)
            FOR tI := 1 TO 8 DO
                IF sK < tN - 2 THEN
                    IF NOT sReturn AND GVL_TestData.X[tA + sK + 1] < tX THEN
                        sK := sK + 1;
                    ELSIF sReturn AND GVL_TestData.X[tA + sK + 1] > tX THEN
                        sK := sK + 1;
                    END_IF;
                END_IF;
            END_FOR;
            tX0 := GVL_TestData.X[tA + sK];
            tX1 := GVL_TestData.X[tA + sK + 1];
            tF0 := GVL_TestData.F[tA + sK];
            tF1 := GVL_TestData.F[tA + sK + 1];
            IF NOT sReturn THEN
                IF tX >= tX1 THEN
                    tF := tF1 + (tX - tX1) * 25.0;
                ELSIF tX <= tX0 OR tX1 - tX0 < 0.000001 THEN
                    tF := tF0;
                ELSE
                    tF := tF0 + (tF1 - tF0) * (tX - tX0) / (tX1 - tX0);
                END_IF;
            ELSE
                IF tX >= tX0 THEN
                    tF := tF0 + (tX - tX0) * 25.0;
                ELSIF tX <= tX1 OR tX0 - tX1 < 0.000001 THEN
                    tF := tF1;
                ELSE
                    tF := tF1 + (tF0 - tF1) * (tX - tX1) / (tX0 - tX1);
                END_IF;
            END_IF;
        END_IF;
    {endregion}

    {region "Outputs"}
        Pos := sPos;
        Force := tF;
        ClampClosed := sClamp >= 0.25;
        ClampOpen := sClamp <= 0.0;
        Moved := sMoved;
    {endregion}
END_FUNCTION_BLOCK

(* ---- PLC_PRG.st ---- *)
// Port of OB1 "Main" with the instance DB "InstTestBench": runs the bench by itself after the start.
PROGRAM PLC_PRG
VAR
    Bench : FB_TestBench;
END_VAR
(* @IMPLEMENTATION *)
Bench();
